(* IEC 61131-3 sources: rusty/compiler/plc_cfc/fixtures/blocks/valid/program_call, 1 file *)

(* ---- counter.st ---- *)
PROGRAM counter
VAR_INPUT
    in : DINT;
END_VAR
VAR_OUTPUT
    out : DINT;
END_VAR
    out := out + in;
END_PROGRAM
